{attribute 'qualified_only'}
{attribute 'strict'}
{attribute 'to_string'}
TYPE L_Apertures :
(
    SL1L0 := 1,
    SL2L0 := 2
);
END_TYPE

(* stored: Version 1.1.0.1
   DUT L_Apertures: Id {81aad000-5d47-45fe-a236-7c80dfbb79b7} *)
